PROGRAM PRG_3_PMPS_POST
VAR
    fbArbiterIO: FB_SubSysToArbiter_IO;
END_VAR

GVL.fbFastFaultOutput1.Execute();
GVL.fbFastFaultOutput2.Execute();

fbArbiterIO(
    Arbiter:=GVL.fbArbiter,
    fbFFHWO:=GVL.fbFastFaultOutput1);

END_PROGRAM

(* stored: Version 1.1.0.1, ProductVersion 3.1.4022.18
   POU PRG_3_PMPS_POST: Id {ae2b5b23-f406-4591-b6ea-00080d408961}, SpecialFunc None *)
